(* IEC 61131-3 sources: kns-pump-station/src/POUs/Log/F_AlarmCode, 2 files *)

(* ---- F_AlarmCode.decl.st ---- *)
// Назначение: код записи журнала по номеру (CSV, DESIGN, раздел 9.2): устройство — <TAG>.<SUFFIX> по
//             GVL_DeviceList (номер = dev_no · 10 + слот, суффиксы слотов — таблица контракта plc-process-lib,
//             раздел 19), станция — KNS1.<SUFFIX> (100000 + slot, 04 §15), LIC101 — LIC101.<SUFFIX> (100100 +
//             слот), событие станции — KNS1.E<код> (101000 + код, 04 §16). Неизвестный номер — его цифры.
// Автор:      kr0nsch
// Версия:     0.1.0
// Документ:   docs/DESIGN.md, раздел 9.2
FUNCTION F_AlarmCode : STRING(GVL_Const.LOG_CODE_LEN)
VAR_INPUT
    udiId : UDINT;                  // номер тревоги или события
END_VAR
VAR
    uiDevNo : UINT;                 // номер устройства
    uiSlot  : UINT;                 // слот тревоги
    uiI     : UINT;                 // индекс GVL_DeviceList
    sSuffix : STRING(GVL_Const.LOG_SUFFIX_LEN);   // суффикс слота
    eType   : PL.E_DeviceType;      // тип устройства
END_VAR
VAR CONSTANT
    ID_PER_DEVICE : UDINT := 10;    // номер тревоги устройства = dev_no · 10 + слот (контракт 20.5)
    STATION_TAG   : STRING(GVL_Const.LOG_SUFFIX_LEN) := 'KNS1';
    PID_TAG       : STRING(GVL_Const.LOG_SUFFIX_LEN) := 'LIC101';
    EVENT_PREFIX  : STRING(GVL_Const.LOG_SUFFIX_LEN) := 'E';
    AI_SUFFIX  : ARRAY[0..GVL_Const.ALM_SLOT_MAX] OF STRING(GVL_Const.LOG_SUFFIX_LEN) :=
        ['HH', 'H', 'L', 'LL', 'FAIL', 'OOR', '', ''];
    DI_SUFFIX  : ARRAY[0..GVL_Const.ALM_SLOT_MAX] OF STRING(GVL_Const.LOG_SUFFIX_LEN) :=
        ['ALM', 'FAIL', '', '', '', '', '', ''];
    MOT_SUFFIX : ARRAY[0..GVL_Const.ALM_SLOT_MAX] OF STRING(GVL_Const.LOG_SUFFIX_LEN) :=
        ['FTS', 'FBL', 'FTP', 'UCR', 'EXT', 'ILK', 'COM', 'SPD'];
    VLV_SUFFIX : ARRAY[0..GVL_Const.ALM_SLOT_MAX] OF STRING(GVL_Const.LOG_SUFFIX_LEN) :=
        ['FTO', 'FTC', 'BLS', 'PLS', 'TRQ', 'EXT', 'ILK', ''];
    CV_SUFFIX  : ARRAY[0..GVL_Const.ALM_SLOT_MAX] OF STRING(GVL_Const.LOG_SUFFIX_LEN) :=
        ['DEV', 'FBF', 'POS', 'ILK', '', '', '', ''];
    PID_SUFFIX : ARRAY[0..GVL_Const.ALM_SLOT_MAX] OF STRING(GVL_Const.LOG_SUFFIX_LEN) :=
        ['PVF', '', '', '', '', '', '', ''];
    // тревоги станции по slot 1…13 (E_StationAlarm, 04 §15)
    STN_SUFFIX : ARRAY[1..GVL_Const.STN_ALARM_COUNT] OF STRING(GVL_Const.LOG_SUFFIX_LEN) :=
        ['EHL', 'DRY', 'LACK', 'NORES', 'ATS', 'FLOAT', 'LDEV', 'STEP', 'NOAUTO', 'UL1', 'UL2', 'UL3', 'SIM'];
END_VAR

(* ---- F_AlarmCode.impl.st ---- *)
F_AlarmCode := UDINT_TO_STRING(udiId);
IF udiId >= GVL_Const.STN_EVENT_ID_BASE THEN
    // событие станции: KNS1.E<код>
    F_AlarmCode := CONCAT(CONCAT(STATION_TAG, '.'),
                          CONCAT(EVENT_PREFIX, UDINT_TO_STRING(udiId - GVL_Const.STN_EVENT_ID_BASE)));
ELSIF udiId >= GVL_Const.LIC101_ALARM_ID_BASE
      AND udiId <= GVL_Const.LIC101_ALARM_ID_BASE + GVL_Const.ALM_SLOT_MAX THEN
    sSuffix := PID_SUFFIX[UDINT_TO_UINT(udiId - GVL_Const.LIC101_ALARM_ID_BASE)];
    IF LEN(sSuffix) > 0 THEN
        F_AlarmCode := CONCAT(CONCAT(PID_TAG, '.'), sSuffix);
    END_IF
ELSIF udiId > GVL_Const.STN_ALARM_ID_BASE AND udiId <= GVL_Const.STN_ALARM_ID_BASE + GVL_Const.STN_ALARM_COUNT THEN
    F_AlarmCode := CONCAT(CONCAT(STATION_TAG, '.'), STN_SUFFIX[UDINT_TO_UINT(udiId - GVL_Const.STN_ALARM_ID_BASE)]);
ELSIF udiId < GVL_Const.STN_ALARM_ID_BASE THEN
    // устройство перечня: dev_no · 10 + слот
    uiDevNo := UDINT_TO_UINT(udiId / ID_PER_DEVICE);
    uiSlot := UDINT_TO_UINT(udiId MOD ID_PER_DEVICE);
    IF uiSlot <= GVL_Const.ALM_SLOT_MAX THEN
        FOR uiI := 1 TO GVL_DeviceList.DEVICE_COUNT DO
            IF GVL_DeviceList.auiDevNo[uiI] = uiDevNo THEN
                eType := GVL_DeviceList.aeDevType[uiI];
                IF eType = PL.E_DeviceType.AnalogInput THEN
                    sSuffix := AI_SUFFIX[uiSlot];
                ELSIF eType = PL.E_DeviceType.DigitalInput THEN
                    sSuffix := DI_SUFFIX[uiSlot];
                ELSIF eType = PL.E_DeviceType.Motor OR eType = PL.E_DeviceType.MotorVfd THEN
                    sSuffix := MOT_SUFFIX[uiSlot];
                ELSIF eType = PL.E_DeviceType.Valve THEN
                    sSuffix := VLV_SUFFIX[uiSlot];
                ELSIF eType = PL.E_DeviceType.ControlValve THEN
                    sSuffix := CV_SUFFIX[uiSlot];
                ELSIF eType = PL.E_DeviceType.Pid THEN
                    sSuffix := PID_SUFFIX[uiSlot];
                ELSE
                    sSuffix := '';
                END_IF
                IF LEN(sSuffix) = 0 THEN
                    sSuffix := UINT_TO_STRING(uiSlot);   // слот без суффикса в контракте — номер слота
                END_IF
                F_AlarmCode := CONCAT(CONCAT(GVL_DeviceList.asTag[uiI], '.'), sSuffix);
                RETURN;
            END_IF
        END_FOR
    END_IF
END_IF
